(* CODESYS project tccamerakeyenceix.library
   Company: TcNexa
   DefaultNamespace: TcNexa_Devices_Camera_TcCameraKeyenceIX
   Version: 1.0.0.0
   Placeholder: TcCameraKeyenceIX
   Author: ATI Software Engineering
   Title: TcCameraKeyenceIX

Project tree, tasks and I/O mapping:
  libraries: Tc2_Standard, 3.4.5.0 (Beckhoff Automation GmbH); Tc2_System, 3.6.4.0 (Beckhoff Automation GmbH); Tc3_Module, 3.4.5.0 (Beckhoff Automation GmbH); TcCamera, 1.0.0.0 (TcNexa); TcDeviceBase, * (TcNexa); TcProcess, 1.0.0.0 (TcNexa)
  DIO/
    function block FB_CameraKeyenceIX_DIO [ST]: inRunMode, overallResult, targetProgramNumber, _handleIO, FB_main, getToolResult, inspect, setProgramNumber
  Tests/
    program PRG_TEST [ST]
*)

// DIO/FB_CameraKeyenceIX_DIO
FUNCTION_BLOCK FB_CameraKeyenceIX_DIO EXTENDS TcNexa_Devices_Base_TcDeviceBase.FB_DeviceBase IMPLEMENTS TcNexa_Devices_Camera_TcCamera.I_Camera
VAR
	IN1					AT %I* : BOOL;
	IN2					AT %I* : BOOL;
	IN3					AT %I* : BOOL;
	IN4					AT %I* : BOOL;
	IN5					AT %I* : BOOL;
	IN6					AT %I* : BOOL;
	IN7					AT %I* : BOOL;
	IN8					AT %I* : BOOL;
	IN9					AT %I* : BOOL;
	IN10				AT %I* : BOOL;
	OUT1				AT %Q* : BOOL;
	OUT2				AT %Q* : BOOL;
	OUT3				AT %Q* : BOOL;
	OUT4				AT %Q* : BOOL;
	OUT5				AT %Q* : BOOL;
	OUT6				AT %Q* : BOOL;
	OUT7				AT %Q* : BOOL;
	OUT8				AT %Q* : BOOL;
	(* IO *)
	_isTotalStatusOk	: BOOL;
	_isBusy				: BOOL;
	_inError			: BOOL;
	_inRunMode			: BOOL;
	_toolResult			: ARRAY[1..6] OF BOOL;
	_trigger			: BOOL;
	_targetProgram		: UINT;
END_VAR

PROPERTY inRunMode : BOOL
GET
inRunMode:= _inRunMode;
END_GET
END_PROPERTY

PROPERTY overallResult : BOOL
GET
overallResult:= _isTotalStatusOk;
END_GET
END_PROPERTY

PROPERTY targetProgramNumber : UINT
GET
targetProgramNumber:= _targetProgram;
END_GET
SET
_targetProgram:= targetProgramNumber;
END_SET
END_PROPERTY

METHOD PROTECTED _handleIO
VAR_INPUT
END_VAR
(* Inputs *)
_isTotalStatusOk:= IN1;
_isBusy:= IN2;
_inError:= IN3;
_inRunMode:= IN4;
_toolResult[1]:= IN5;
_toolResult[2]:= IN6;
_toolResult[3]:= IN7;
_toolResult[4]:= IN8;
_toolResult[5]:= IN9;
_toolResult[6]:= IN10;

(* Outputs *)
OUT1:= _trigger;
OUT2:= _targetProgram.0;
OUT3:= _targetProgram.1;
OUT4:= _targetProgram.2;
OUT5:= _targetProgram.3;
OUT6:= _targetProgram.4;
END_METHOD

METHOD FB_main
VAR_INPUT
END_VAR
SUPER^.FB_main();

_handleIO();
END_METHOD

METHOD PUBLIC getToolResult : BOOL
VAR_INPUT
	index			: UINT;
	Response		: REFERENCE TO TcNexa_Components_TcProcess.FB_MethodResponse;
END_VAR
IF (index < 1) OR (index > 6) THEN
	IF __ISVALIDREF(Response) THEN Response.setFail(description:= 'Invalid index'); END_IF
ELSE
	getToolResult:= _toolResult[index];
	IF __ISVALIDREF(Response) THEN Response.setPass(); END_IF
END_IF
END_METHOD

METHOD inspect
VAR_INPUT
	Response	: REFERENCE TO TcNexa_Devices_Camera_TcCamera.TcNexa_Components_TcProcess.FB_MethodResponse;
END_VAR
_methodState:= _methodHeader(methodName:= 'inspect');

IF _methodState.init THEN
	IF NOT _inRunMode THEN
		_InternalResponse.setFail(
			description:= Tc2_Standard.CONCAT(
				STR1:= _nameTag, 
				STR2:= ' is not in run'));
	ELSIF _inError THEN
		_InternalResponse.setFail(
			description:= Tc2_Standard.CONCAT(
				STR1:= _nameTag, 
				STR2:= ' is in error'));
	END_IF
	_trigger:= FALSE;
ELSIF _methodState.execute THEN	
	CASE _Step.actual OF
		0:	
			_trigger:= TRUE;
			IF _isBusy THEN
				_Step.inc();
			END_IF
		1:
			IF _inError THEN
				_InternalResponse.setFail(
					description:= Tc2_Standard.CONCAT(
						STR1:= _nameTag, 
						STR2:= ' is in error'));
			ELSIF _isBusy THEN
				_InternalResponse.setBusy(
					description:= _getBusyDescription(
						description:= 'in progress'));
			ELSE
				_InternalResponse.setPass();
			END_IF
	END_CASE
END_IF

IF NOT _InternalResponse.busy THEN
	_trigger:= FALSE;
END_IF

_methodFooter(Response:= Response);
END_METHOD

METHOD setProgramNumber
VAR_INPUT
	programNumber	: UINT;
	Response	: REFERENCE TO TcNexa_Devices_Camera_TcCamera.TcNexa_Components_TcProcess.FB_MethodResponse;
END_VAR
_methodState:= _methodHeader(methodName:= 'setProgramNumber');

_targetProgram:= programNumber;
_InternalResponse.setPass();

_methodFooter(Response:= Response);
END_METHOD

END_FUNCTION_BLOCK

// Tests/PRG_TEST
PROGRAM PRG_TEST
VAR
END_VAR

END_PROGRAM
